(* PLC project , Example Fixture *)

PROGRAM Main
  VAR_OUTPUT
    Run : BOOL;
  END_VAR

(* LD diagram, written out as Structured Text *)
Run := %IX0.3;
END_PROGRAM

CONFIGURATION c
  RESOURCE r ON PLC
  END_RESOURCE
END_CONFIGURATION
